// TIA Portal V21 export
// export: Created 2026-11-07T15:50:49.9861994Z, ExportSetting WithDefaults, DisplayName Totally Integrated Automation Portal, DisplayVersion V21, DisplayName STEP 7 Professional, DisplayVersion V21, DisplayName STEP 7 Safety, DisplayVersion V21, DisplayName Tech WebApplication, DisplayVersion V21, DisplayName WinCC Basic/Comfort/Advanced, DisplayVersion V21, DisplayName WinCC Unified, DisplayVersion V21
Screen "R04_BtnInv"  1024x768, Number=43, Template=Tpl
  ScreenLayer 
    Button "P_BtnInv" at 10,10 size 100x30  Mode=Text, StyleItem=Button, TextOff="BTN", TextOn="BTN"
      on Press: InvertBit(Tag := P_SwOn)
